TYPE ET_Gr02Manual :
(
	ET_Gr02Manual_eWaitExecute := 0,
	ET_Gr02Manual_eSetPosAxis5,
	ET_Gr02Manual_eWfSetPosAxis5,
	ET_Gr02Manual_eCouplingAxis1_4,
	ET_Gr02Manual_eWfCouplingAxis1_4,
	ET_Gr02Manual_eDone := 197,
	ET_Gr02Manual_eError := 198,
	ET_Gr02Manual_eNoExecute := 199
);
END_TYPE

(* stored: Version 1.1.0.1, ProductVersion 3.1.4024.15
   DUT ET_Gr02Manual: Id {eb2e9b55-f8a8-4c4c-95f6-7c384d3689c7} *)
